Fanuc KAREL source: KT00077.KL

PROGRAM KT00077
%NOLOCKGROUP
VAR
  R1: REAL
  Y2: ARRAY[2] OF BYTE
  OUT: INTEGER
BEGIN
  R1 = 2.0
    Y2[1] = 3
  OUT = R1 * Y2[1]
END KT00077
